// TIA Portal V21 export
// export: Created 2026-08-21T20:18:45.5439062Z, ExportSetting None, DisplayName Totally Integrated Automation Portal, DisplayVersion V21, DisplayName STEP 7 Professional, DisplayVersion V21, DisplayName STEP 7 Safety, DisplayVersion V21, DisplayName Tech WebApplication, DisplayVersion V21, DisplayName WinCC Basic/Comfort/Advanced, DisplayVersion V21, DisplayName WinCC Professional, DisplayVersion V21, DisplayName WinCC Unified, DisplayVersion V21
DATA_BLOCK "ModuleTypePackageRevision"   // DB59
TITLE = ModuleTypePackageRevision
{ S7_Optimized_Access := 'TRUE' }
AUTHOR : Siemens AG
FAMILY : MTP
VERSION : 1.0
// The version information of the entire MTP
// stored: InstanceOfName typeMTPModuleTypePackageRevision, InstanceOfType UDT
"typeMTPModuleTypePackageRevision"
   // VAR
   //    ModuleTypePackageRevision { ExternalAccessible := 'False'; ExternalVisible := 'False'; ExternalWritable := 'False'} : String := '3.0.0';
   // END_VAR
BEGIN
END_DATA_BLOCK
